Fanuc KAREL source: KT00596.KL

PROGRAM KT00596
%NOLOCKGROUP
VAR
  R1: REAL
  I2: INTEGER
  OUT: STRING[80]
BEGIN
  R1 = 2.0
    I2 = 3
  OUT = R1 + I2
END KT00596
